// TIA Portal V21 export
FUNCTION_BLOCK "FB_AnaTimerInIf"   // FB11, SCL
TITLE = Analyzer: timer called inside IF
{ S7_Optimized_Access := 'TRUE' }
// Rule C26a: the timer is only called while Enable is TRUE, so it freezes otherwise
// stored: MemoryReserve 100, SetENOAutomatically false
   VAR_INPUT
      Enable : Bool;   // Enable
      Start : Bool;   // Timer input
   END_VAR
   VAR_OUTPUT
      Done : Bool;   // Timer output
   END_VAR
   VAR
      Delay { S7_SetPoint := 'True'} : TON_TIME;   // On-delay timer
   END_VAR
BEGIN

       IF #Enable THEN
           #Delay(IN := #Start, PT := T#1s);
       END_IF;
       #Done := #Delay.Q;
END_FUNCTION_BLOCK
